TYPE "ST_DeclarationLeafHal"
VERSION : 0.1
   STRUCT
      Sample : DInt;
      Permit : Bool := TRUE;
      Finish : Bool;
      BackgroundFault : Bool;
      Diag : "ST_Diagnostic";
      LaterDiag : "ST_Diagnostic";
      ExitHold : Bool;
      Verdict : DInt := 1;
   END_STRUCT;

END_TYPE

